FUNCTION_BLOCK Level_Control (* Composite Function Block Type *)
  (* Standard: 61499-2 *)
  (* Version 0.0, 1/6/2020, prana, nxtControl GmbH, template *)
  PACKAGE Main;
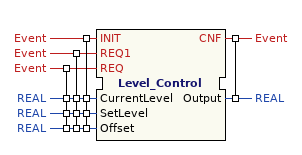
  EVENT_INPUT
    INIT WITH CurrentLevel, SetLevel, Offset; (* Initialization Request *)
    REQ1 WITH CurrentLevel, SetLevel, Offset;
    REQ WITH CurrentLevel, SetLevel, Offset;
  END_EVENT
  EVENT_OUTPUT
    CNF WITH Output; (* Execution Confirmation *)
  END_EVENT
  VAR_INPUT
    CurrentLevel : REAL; (* Input event qualifier *)
    SetLevel : REAL;
    Offset : REAL;
  END_VAR
  VAR_OUTPUT
    Output : REAL; (* Output event qualifier *)
  END_VAR
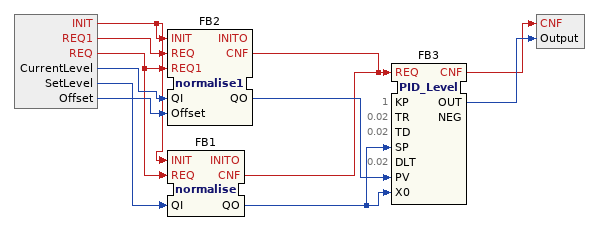
  FBS
    FB1 : normalise;
    FB2 : normalise1;
    FB3 : PID_Level(KP := 1, TR := 0.02, TD := 0.02, DLT := 0.02);
  END_FBS
  EVENT_CONNECTIONS
    INIT TO FB2.INIT;
    FB1.CNF TO FB3.REQ;
    FB2.CNF TO FB3.REQ;
    FB3.CNF TO CNF;
    INIT TO FB1.INIT;
    REQ1 TO FB2.REQ;
    REQ TO FB1.REQ;
    REQ TO FB2.REQ1;
  END_CONNECTIONS
  DATA_CONNECTIONS
    SetLevel TO FB1.QI;
    CurrentLevel TO FB2.QI;
    FB1.QO TO FB3.X0;
    FB1.QO TO FB3.SP;
    FB2.QO TO FB3.PV;
    FB3.OUT TO Output;
    Offset TO FB2.Offset;
  END_CONNECTIONS
END_FUNCTION_BLOCK
